(* IEC 61131-3 sources: SemantiST/compiler/intake/normalize/probes/standard-formal-arguments, 2 files *)

(* ---- original.st ---- *)
FUNCTION main : DINT
printf('%d %d$N', MIN(IN1 := 3, IN2 := 9), LIMIT(MN := 0, IN := 12, MX := 7));
main := 0;
END_FUNCTION

(* ---- rewritten.st ---- *)
FUNCTION main : DINT
printf('%d %d$N', MIN(3, 9), LIMIT(0, 12, 7));
main := 0;
END_FUNCTION
